SUBAPPLICATION logiBUS_AI_Raw_VT_AR_Param_OPC (* Wie logiBUS_AI_Raw_VT_AR_OPC, aber Hysterese, TimeDelta und TimeRateLimit des AI einstellbar (INI + Web), Wirkung nach Neustart *)
  (* Standard: 61499-2; Description: Copyright (c) 2026 Meisterschulen am Ostbahnhof This program and the accompanying materials are made available under the terms of the Eclipse Public License 2.0 which is available at https://www.eclipse.org/legal/epl-2.0/ SPDX-License-Identifier: EPL-2.0 *)
  (* Version 1.0, 2026-10-30, Franz Höpfinger, Meisterschulen am Ostbahnhof, Kopie von logiBUS_AI_Raw_VT_AR_OPC. Franz: Achslenkung pendelt beim Zentrieren - Hysterese 50 Digits (~9 %) groesser als das Null-Fenster +-2 % (~21 Digits). AnalogInput_hysteresis/TimeDelta/TimeRateLimit jetzt je OPC_TO_AR2_OUT (Web) + INI_AR2 (Keys AI_Hysterese/AI_TimeDelta/AI_TimeRateLimit in sSection), Defaults per Parameter. Werden vor logiBUS_AI_IDA.INIT geladen, eine Aenderung wirkt erst nach Neustart (wie FilterTimeS). INIT-Kette AI -> Q_NumericValue_RAW -> AR_PUBLISH_RAW wie im Original (Franz, 2026-10-30). VT-Rohwertanzeige per AUDI_D_FF_TMIN (500 ms) gedrosselt, AR_OUT/Publish ungedrosselt (Franz: Regelung schnell, Anzeige darf hinterherhinken). Siehe KALIBRIERUNG_Achslenkung_Winkel.md. *)
  PACKAGE MyLib::sys;
  IMPORT logiBUS::io::AI::logiBUS_AI;
  IMPORT logiBUS::io::AI::logiBUS_AI_S;
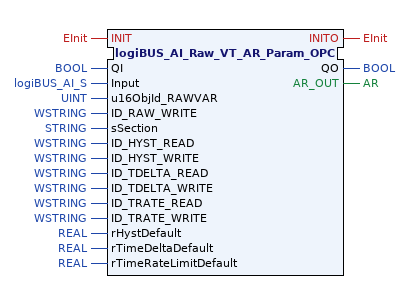
  EVENT_INPUT
    INIT : EInit; (* Initialization Request *)
  END_EVENT
  EVENT_OUTPUT
    INITO : EInit; (* Initialization Confirm *)
  END_EVENT
  VAR_INPUT
    QI : BOOL := TRUE; (* Quality Input - TRUE to enable service *)
    Input : logiBUS::io::AI::logiBUS_AI_S := logiBUS_AI::Invalid; (* Identify the Input AnalogInput_I1..I8 *)
    u16ObjId_RAWVAR : UINT; (* Object ID CNumberVariable (Rohwert 0-4095, unkalibriert, reine Diagnose-Anzeige) *)
    ID_RAW_WRITE : WSTRING; (* Rohwert-Ruckmelde-Adresse (REAL 0-4095, ACTION=PUBLISH) *)
    sSection : STRING; (* INI-Section (gleich wie Kalibrierung) *)
    ID_HYST_READ : WSTRING; (* Web-Override Hysterese (Digits) *)
    ID_HYST_WRITE : WSTRING; (* Rueckmeldung Hysterese (Digits) *)
    ID_TDELTA_READ : WSTRING; (* Web-Override TimeDelta (ms) *)
    ID_TDELTA_WRITE : WSTRING; (* Rueckmeldung TimeDelta (ms) *)
    ID_TRATE_READ : WSTRING; (* Web-Override TimeRateLimit (ms) *)
    ID_TRATE_WRITE : WSTRING; (* Rueckmeldung TimeRateLimit (ms) *)
    rHystDefault : REAL := 3.0; (* Default Hysterese (Digits) *)
    rTimeDeltaDefault : REAL := 100.0; (* Default TimeDelta (ms) *)
    rTimeRateLimitDefault : REAL := 20.0; (* Default TimeRateLimit (ms) *)
  END_VAR
  VAR_OUTPUT
    QO : BOOL; (* Quality Output - TRUE if service executed successfully *)
  END_VAR
  PLUGS
    AR_OUT : adapter::types::unidirectional::AR; (* Rohwert als AR, fertig fuer CALIBRATE.X *)
  END_PLUGS
  FBS
    logiBUS_AI_IDA : logiBUS::io::AI::logiBUS_AI_IDA;
    INI_Hyst : eclipse4diac::storage::INI_AR2(SETM := TRUE, KEY := 'AI_Hysterese');
    ToAD_Hyst : adapter::conversion::unidirectional::AR_TO_AD_NUM;
    ToDWORD_Hyst : adapter::conversion::unidirectional::AD_D_TO_DWORD;
    INI_TDelta : eclipse4diac::storage::INI_AR2(SETM := TRUE, KEY := 'AI_TimeDelta');
    ToAD_TDelta : adapter::conversion::unidirectional::AR_TO_AD_NUM;
    ToDWORD_TDelta : adapter::conversion::unidirectional::AD_D_TO_DWORD;
    INI_TRate : eclipse4diac::storage::INI_AR2(SETM := TRUE, KEY := 'AI_TimeRateLimit');
    ToAD_TRate : adapter::conversion::unidirectional::AR_TO_AD_NUM;
    ToDWORD_TRate : adapter::conversion::unidirectional::AD_D_TO_DWORD;
    AD_TO_AUDI : adapter::conversion::unidirectional::AD_TO_AUDI;
    AUDI_SPLIT_2 : adapter::events::unidirectional::AUDI_SPLIT_2;
    RateLimit_Anzeige : adapter::events::unidirectional::AUDI_D_FF_TMIN(Tmin := T#500ms); (* Nur VT-Anzeige gedrosselt, AR_OUT (Regelung) ungedrosselt *)
    Q_NumericValue_RAW : isobus::UT::Q::Q_NumericValue_AUDI;
    AUDI_TO_AR : adapter::conversion::unidirectional::AUDI_TO_AR;
    AR_SPLIT_2_Raw : adapter::events::unidirectional::AR_SPLIT_2;
    AR_PUBLISH_RAW : adapter::net::AR_PUBLISH_1;
    AND_QO : iec61131::booleanOperators::AND_BOOL_3;
  END_FBS
  SUBAPPS
    Par_Hyst : MyLib::sys::OPC_TO_AR2_OUT;
    Par_TDelta : MyLib::sys::OPC_TO_AR2_OUT;
    Par_TRate : MyLib::sys::OPC_TO_AR2_OUT;
  END_SUBAPPS
  EVENT_CONNECTIONS
    logiBUS_AI_IDA.INITO TO Q_NumericValue_RAW.INIT;
    Q_NumericValue_RAW.INITO TO AR_PUBLISH_RAW.INIT;
    AR_PUBLISH_RAW.INITO TO INITO;
    AR_PUBLISH_RAW.INITO TO AND_QO.REQ;
    INIT TO Par_TRate.INIT;
    Par_TRate.INITO TO INI_TRate.INIT;
    INI_TRate.INITO TO Par_TDelta.INIT;
    Par_TDelta.INITO TO INI_TDelta.INIT;
    INI_TDelta.INITO TO Par_Hyst.INIT;
    Par_Hyst.INITO TO INI_Hyst.INIT;
    INI_Hyst.INITO TO logiBUS_AI_IDA.INIT;
  END_CONNECTIONS
  DATA_CONNECTIONS
    Input TO logiBUS_AI_IDA.Input;
    u16ObjId_RAWVAR TO Q_NumericValue_RAW.u16ObjId;
    ID_RAW_WRITE TO AR_PUBLISH_RAW.ID;
    QI TO Q_NumericValue_RAW.QI;
    QI TO logiBUS_AI_IDA.QI;
    QI TO AR_PUBLISH_RAW.QI;
    Q_NumericValue_RAW.QO TO AND_QO.IN1;
    logiBUS_AI_IDA.QO TO AND_QO.IN2;
    AR_PUBLISH_RAW.QO TO AND_QO.IN3;
    AND_QO.OUT TO QO;
    rHystDefault TO INI_Hyst.DEFAULT_VALUE;
    sSection TO INI_Hyst.SECTION;
    QI TO INI_Hyst.QI;
    QI TO Par_Hyst.QI;
    ID_HYST_READ TO Par_Hyst.ID_READ;
    ID_HYST_WRITE TO Par_Hyst.ID_WRITE;
    ToDWORD_Hyst.IN TO logiBUS_AI_IDA.AnalogInput_hysteresis;
    rTimeDeltaDefault TO INI_TDelta.DEFAULT_VALUE;
    sSection TO INI_TDelta.SECTION;
    QI TO INI_TDelta.QI;
    QI TO Par_TDelta.QI;
    ID_TDELTA_READ TO Par_TDelta.ID_READ;
    ID_TDELTA_WRITE TO Par_TDelta.ID_WRITE;
    ToDWORD_TDelta.IN TO logiBUS_AI_IDA.TimeDelta;
    rTimeRateLimitDefault TO INI_TRate.DEFAULT_VALUE;
    sSection TO INI_TRate.SECTION;
    QI TO INI_TRate.QI;
    QI TO Par_TRate.QI;
    ID_TRATE_READ TO Par_TRate.ID_READ;
    ID_TRATE_WRITE TO Par_TRate.ID_WRITE;
    ToDWORD_TRate.IN TO logiBUS_AI_IDA.TimeRateLimit;
  END_CONNECTIONS
  ADAPTER_CONNECTIONS
    logiBUS_AI_IDA.IN TO AD_TO_AUDI.AD_IN;
    AD_TO_AUDI.AUDI_OUT TO AUDI_SPLIT_2.IN;
    AUDI_SPLIT_2.OUT1 TO RateLimit_Anzeige.I;
    RateLimit_Anzeige.Q TO Q_NumericValue_RAW.u32NewValue;
    AUDI_SPLIT_2.OUT2 TO AUDI_TO_AR.AUDI_IN;
    AUDI_TO_AR.AR_OUT TO AR_SPLIT_2_Raw.IN;
    AR_SPLIT_2_Raw.OUT1 TO AR_OUT;
    AR_SPLIT_2_Raw.OUT2 TO AR_PUBLISH_RAW.IN;
    Par_Hyst.VALUEO TO INI_Hyst.VAL;
    Par_Hyst.VALUE_OUT TO ToAD_Hyst.AR_IN;
    ToAD_Hyst.AD_OUT TO ToDWORD_Hyst.AD_IN;
    Par_TDelta.VALUEO TO INI_TDelta.VAL;
    Par_TDelta.VALUE_OUT TO ToAD_TDelta.AR_IN;
    ToAD_TDelta.AD_OUT TO ToDWORD_TDelta.AD_IN;
    Par_TRate.VALUEO TO INI_TRate.VAL;
    Par_TRate.VALUE_OUT TO ToAD_TRate.AR_IN;
    ToAD_TRate.AD_OUT TO ToDWORD_TRate.AD_IN;
  END_CONNECTIONS
END_SUBAPPLICATION
